(* IEC 61131-3 sources: linesight/plc/src, 5 files *)

(* ---- E_PackML.st ---- *)
// DUT (Enumeration). Numery stanów zgodne z PackML (ISA-TR88.00.02, PackTag Status.StateCurrent).
// Podzbiór: bez stanów przejściowych Holding/Unholding/Suspending/Unsuspending i bez Completing/Complete.
{attribute 'qualified_only'}
TYPE E_PackML :
(
    Clearing  := 1,
    Stopped   := 2,
    Starting  := 3,
    Idle      := 4,
    Suspended := 5,   // przyczyna zewnętrzna: brak produktu na wejściu
    Execute   := 6,
    Stopping  := 7,
    Aborting  := 8,
    Aborted   := 9,
    Held      := 11,  // przyczyna wewnętrzna: zator w maszynie
    Resetting := 15
) INT;
END_TYPE

(* ---- GVL_Line.st ---- *)
// GVL: interfejs linii – wszystko, co wystawiamy przez OPC UA (E3-04).
{attribute 'qualified_only'}
VAR_GLOBAL
    // --- Komendy operatora (zbocze narastające; odpowiednik PackTag Command.CntrlCmd) ---
    xCmdReset     : BOOL;   // Stopped -> Resetting -> Idle
    xCmdStart     : BOOL;   // Idle -> Starting -> Execute
    xCmdStop      : BOOL;   // Idle/Execute/Held/Suspended -> Stopping -> Stopped
    xCmdAbort     : BOOL;   // dowolny stan -> Aborting -> Aborted (wyłącznik awaryjny)
    xCmdClear     : BOOL;   // Aborted -> Clearing -> Stopped

    // --- Wstrzykiwanie awarii (poziom: TRUE = usterka trwa) ---
    xInjJam       : BOOL;   // zator                 -> Held,      iStopReason 101
    xInjNoProduct : BOOL;   // brak produktu         -> Suspended, iStopReason 201
    xInjFault     : BOOL;   // awaria (np. napęd)    -> Aborted,   iStopReason 301
    xInjSlow      : BOOL;   // degradacja: czas cyklu +40 % (dane do wykrywania anomalii, etap 4)
    xInjWear      : BOOL;   // E4-06: zużycie napędu (łożysko) narasta przez tWearRamp; FALSE = naprawa

    // --- Nastawy ---
    tCycleNominal : TIME := T#1500MS;   // nominalny czas cyklu (1 sztuka)
    tWearRamp     : TIME := T#20M;      // E4-06: czas narastania zużycia napędu do 100 %

    // --- Status (tylko do odczytu dla świata) ---
    iStateCurrent    : INT;     // Status.StateCurrent (numer stanu PackML)
    iStopReason      : INT;     // Admin.StopReason.ID: 0 brak, 1 stop operatora, 101 zator,
                                // 201 brak produktu, 301 awaria, 302 abort operatora
    udiProdProcessed : UDINT;   // Admin.ProdProcessedCount (licznik narastający, nie kasujemy)
    udiCycleTime_ms  : UDINT;   // czas ostatniego cyklu [ms] (symulowany)
    rMachSpeed       : REAL;    // Status.CurMachSpeed [szt./min], 0 poza Execute

    // --- E4-06: napęd taśmy (FB_DriveSim), wartości na sztukę ---
    rTorqueMean_Nm   : REAL;    // średni moment w cyklu
    rTorquePeak_Nm   : REAL;    // szczytowy moment w cyklu
    rCurrent_A       : REAL;    // prąd silnika
    rMotorTemp_C     : REAL;    // temperatura silnika (0,1 °C)
    rSimWear         : REAL;    // zużycie 0..1 – prawda symulacji, tylko do oceny modelu (zaokr. 0,01)
END_VAR

(* ---- F_Gauss.st ---- *)
// FUNCTION F_Gauss – szum o rozkładzie zbliżonym do normalnego (średnia 0, odchylenie 1).
// Suma 4 liczb równomiernych z LCG (centralne twierdzenie graniczne); wystarcza do symulacji pomiaru.
// Ziarno przekazywane przez VAR_IN_OUT – stan generatora trzyma wywołujący blok.
// --- część deklaracji ---
FUNCTION F_Gauss : REAL
VAR_IN_OUT
    udiSeed : UDINT;
END_VAR
VAR
    i : INT;
    rSum : REAL;                     // zmienne funkcji startują od 0 przy każdym wywołaniu; nie „s”: S i R to słowa kluczowe IEC (Set/Reset)
END_VAR

// --- część implementacji ---
FOR i := 1 TO 4 DO
    udiSeed := udiSeed * 1103515245 + 12345;
    rSum := rSum + UDINT_TO_REAL((udiSeed / 65536) MOD 32768) / 32768.0;
END_FOR
F_Gauss := (rSum - 2.0) * 1.7320508;    // suma 4 x U(0,1): średnia 2, wariancja 4/12 -> skalowanie do odchylenia 1

(* ---- FB_DriveSim.st ---- *)
// FUNCTION_BLOCK FB_DriveSim – symulacja napędu taśmy (E4-06): moment, prąd, temperatura, zużycie.
// Wartości na sztukę (jak napęd raportujący parametry cyklu), temperatura liczona ciągle.
//   Moment średni   Tm = 2,0 Nm x (1 + 0,15 x zużycie + zimno) + szum 0,06 Nm x (1 + 1,5 x zużycie)
//                   zimno = 0,12 x (40 °C - T) / 18 °C, w zakresie 0..0,12: zimny smar = większe tarcie,
//                   po każdym dłuższym postoju moment jest wyższy o do 12 % i spada, gdy silnik się nagrzeje
//   Moment szczyt.  Tp = Tm x (1,6 + 0,25 x zużycie)     + szum 0,08 Nm x (1 + 2,0 x zużycie)
//   Prąd            I  = 0,8 A + 1,2 A/Nm x Tm            + szum 0,02 A
//   Temperatura     dT/dt = (22 °C + 2,25 x I^2 - T) / 600 s   (inercja 1. rzędu; I = 0 poza Execute)
// Zużycie (np. łożysko): przy xWear rośnie liniowo 0 -> 1 w czasie tWearRamp, bez xWear = 0 (po naprawie).
// Wczesne zużycie ginie w szumie pojedynczej sztuki, a próg na samym momencie myli zużycie z zimnym startem –
// model, który zna temperaturę i kształt cyklu (szczyt/średnia, rozrzut), ma je odróżnić.
// --- część deklaracji ---
FUNCTION_BLOCK FB_DriveSim
VAR_INPUT
    xRun       : BOOL;                 // linia w Execute (napęd pracuje)
    xCycleDone : BOOL;                 // impuls: koniec sztuki – nowe wartości momentu i prądu
    xWear      : BOOL;                 // wstrzyknięte zużycie
    tWearRamp  : TIME := T#20M;        // czas narastania zużycia do 100 %
END_VAR
VAR_OUTPUT
    rTorqueMean : REAL;                // [Nm]
    rTorquePeak : REAL;                // [Nm]
    rCurrent    : REAL;                // [A]
    rTemp       : REAL := 22.0;        // [°C], zaokrąglone do 0,1 (mniej wiadomości przez OPC UA)
    rWear       : REAL;                // 0..1, prawda symulacji – tylko do oceny modelu
END_VAR
VAR
    udiSeed : UDINT := 987654321;
    tLast   : TIME;
    xInit   : BOOL;
    rDt     : REAL;                    // [s] od poprzedniego wywołania
    rT      : REAL := 22.0;            // temperatura bez zaokrąglenia
    rI      : REAL;
    rTm     : REAL;
    rCold   : REAL;                    // dodatkowe tarcie zimnego napędu, 0..0,12
END_VAR
VAR CONSTANT
    T0     : REAL := 2.0;
    TAMB   : REAL := 22.0;
    K_HEAT : REAL := 2.25;
    TAU_S  : REAL := 600.0;
END_VAR

// --- część implementacji ---
IF NOT xInit THEN
    tLast := TIME();
    xInit := TRUE;
END_IF
rDt := TIME_TO_REAL(TIME() - tLast) / 1000.0;
tLast := TIME();

// zużycie
IF xWear AND tWearRamp > T#0S THEN
    rWear := MIN(1.0, rWear + rDt / (TIME_TO_REAL(tWearRamp) / 1000.0));
ELSE
    rWear := 0.0;
END_IF

// temperatura: inercja pierwszego rzędu (metoda Eulera), grzanie proporcjonalne do I^2
IF xRun THEN rI := rCurrent; ELSE rI := 0.0; END_IF
rT := rT + rDt / TAU_S * (TAMB + K_HEAT * rI * rI - rT);
rTemp := DINT_TO_REAL(TRUNC(rT * 10.0)) / 10.0;

// parametry sztuki
IF xCycleDone THEN
    rCold := LIMIT(0.0, 0.12 * (40.0 - rT) / 18.0, 0.12);
    rTm := T0 * (1.0 + 0.15 * rWear + rCold) + 0.06 * (1.0 + 1.5 * rWear) * F_Gauss(udiSeed);
    rTorqueMean := DINT_TO_REAL(TRUNC(rTm * 1000.0)) / 1000.0;
    rTorquePeak := DINT_TO_REAL(TRUNC((rTm * (1.6 + 0.25 * rWear)
                   + 0.08 * (1.0 + 2.0 * rWear) * F_Gauss(udiSeed)) * 1000.0)) / 1000.0;
    rCurrent := DINT_TO_REAL(TRUNC((0.8 + 1.2 * rTm + 0.02 * F_Gauss(udiSeed)) * 1000.0)) / 1000.0;
END_IF

(* ---- PLC_PRG.st ---- *)
// PROGRAM PLC_PRG – maszyna stanów PackML (podzbiór) + symulacja produkcji.
// --- część deklaracji ---
PROGRAM PLC_PRG
VAR
    eState    : E_PackML := E_PackML.Stopped;
    ePrev     : E_PackML := E_PackML.Stopped;
    xNewState : BOOL;
    tonAct    : TON;                 // czas trwania stanów przejściowych (Starting, Stopping, ...)
    tonCycle  : TON;                 // czas cyklu jednej sztuki
    rtReset, rtStart, rtStop, rtAbort, rtClear : R_TRIG;
    tCycle    : TIME := T#1500MS;    // czas bieżącego cyklu (nominalny ± rozrzut)
    udiBase   : UDINT;
    udiSeed   : UDINT := 12345;      // generator pseudolosowy (LCG) do rozrzutu czasu cyklu
    xRun, xRunPrev : BOOL;
    tStart, tNow   : TIME;           // TIME() = czas od startu sterownika; z niego mierzymy rzeczywisty cykl
    xPiece    : BOOL;                // E4-06: impuls – w tym cyklu zadania skończyła się sztuka
    fbDrive   : FB_DriveSim;         // E4-06: symulacja napędu taśmy
END_VAR
VAR CONSTANT
    T_ACT : TIME := T#1S;            // ile trwa każdy stan przejściowy
END_VAR

// --- część implementacji ---
rtReset(CLK := GVL_Line.xCmdReset);
rtStart(CLK := GVL_Line.xCmdStart);
rtStop(CLK := GVL_Line.xCmdStop);
rtAbort(CLK := GVL_Line.xCmdAbort);
rtClear(CLK := GVL_Line.xCmdClear);

// Zegar stanu przejściowego: zeruje się w cyklu, w którym stan się zmienił
xNewState := eState <> ePrev;
ePrev := eState;
tonAct(IN := NOT xNewState, PT := T_ACT);

// Abort ma pierwszeństwo przed wszystkim (jak w PackML: z każdego stanu)
IF (rtAbort.Q OR GVL_Line.xInjFault)
   AND eState <> E_PackML.Aborting AND eState <> E_PackML.Aborted AND eState <> E_PackML.Clearing THEN
    IF GVL_Line.xInjFault THEN
        GVL_Line.iStopReason := 301;
    ELSE
        GVL_Line.iStopReason := 302;
    END_IF
    eState := E_PackML.Aborting;
// Stop operatora z każdego stanu „roboczego”
ELSIF rtStop.Q AND (eState = E_PackML.Idle OR eState = E_PackML.Execute
                    OR eState = E_PackML.Held OR eState = E_PackML.Suspended) THEN
    GVL_Line.iStopReason := 1;
    eState := E_PackML.Stopping;
ELSE
    CASE eState OF
        E_PackML.Stopped:
            IF rtReset.Q THEN eState := E_PackML.Resetting; END_IF

        E_PackML.Resetting:
            GVL_Line.iStopReason := 0;
            IF tonAct.Q THEN eState := E_PackML.Idle; END_IF

        E_PackML.Idle:
            IF rtStart.Q THEN eState := E_PackML.Starting; END_IF

        E_PackML.Starting:
            IF tonAct.Q THEN eState := E_PackML.Execute; END_IF

        E_PackML.Execute:
            IF GVL_Line.xInjJam THEN
                GVL_Line.iStopReason := 101;
                eState := E_PackML.Held;
            ELSIF GVL_Line.xInjNoProduct THEN
                GVL_Line.iStopReason := 201;
                eState := E_PackML.Suspended;
            END_IF

        E_PackML.Held:        // zator usunięty -> wracamy do pracy
            IF NOT GVL_Line.xInjJam THEN
                GVL_Line.iStopReason := 0;
                eState := E_PackML.Execute;
            END_IF

        E_PackML.Suspended:   // produkt wrócił -> wracamy do pracy
            IF NOT GVL_Line.xInjNoProduct THEN
                GVL_Line.iStopReason := 0;
                eState := E_PackML.Execute;
            END_IF

        E_PackML.Stopping:
            IF tonAct.Q THEN eState := E_PackML.Stopped; END_IF

        E_PackML.Aborting:
            IF tonAct.Q THEN eState := E_PackML.Aborted; END_IF

        E_PackML.Aborted:     // kasowanie możliwe dopiero po usunięciu awarii
            IF rtClear.Q AND NOT GVL_Line.xInjFault THEN eState := E_PackML.Clearing; END_IF

        E_PackML.Clearing:
            IF tonAct.Q THEN
                GVL_Line.iStopReason := 0;
                eState := E_PackML.Stopped;
            END_IF
    END_CASE
END_IF

// --- Symulacja produkcji: w Execute jedna sztuka co tCycle ---
// udiCycleTime_ms to ZMIERZONY czas od poprzedniej sztuki (TIME()), a nie zadany tCycle:
// timer widzi czas tylko co cykl zadania, więc rzeczywisty cykl jest dłuższy od zadanego.
xRun := eState = E_PackML.Execute;
IF xRun AND NOT xRunPrev THEN
    tStart := TIME();                // wejście w Execute: liczymy od nowa (postój nie wlicza się do cyklu)
END_IF
xRunPrev := xRun;
tonCycle(IN := xRun, PT := tCycle);
xPiece := tonCycle.Q;
IF tonCycle.Q THEN
    tNow := TIME();
    GVL_Line.udiProdProcessed := GVL_Line.udiProdProcessed + 1;
    GVL_Line.udiCycleTime_ms := TIME_TO_UDINT(tNow - tStart);
    tStart := tNow;
    tonCycle(IN := FALSE);           // kasowanie timera; nowy cykl rusza w następnym cyklu zadania

    // czas następnego cyklu: nominalny (x1,4 przy degradacji) z rozrzutem ±100 ms
    udiBase := TIME_TO_UDINT(GVL_Line.tCycleNominal);
    IF GVL_Line.xInjSlow THEN udiBase := udiBase * 14 / 10; END_IF
    IF udiBase < 300 THEN udiBase := 300; END_IF
    udiSeed := udiSeed * 1103515245 + 12345;
    tCycle := UDINT_TO_TIME(udiBase + (udiSeed / 65536) MOD 201 - 100);
END_IF

// --- E4-06: napęd taśmy ---
fbDrive(xRun := xRun, xCycleDone := xPiece, xWear := GVL_Line.xInjWear, tWearRamp := GVL_Line.tWearRamp);
GVL_Line.rTorqueMean_Nm := fbDrive.rTorqueMean;
GVL_Line.rTorquePeak_Nm := fbDrive.rTorquePeak;
GVL_Line.rCurrent_A     := fbDrive.rCurrent;
GVL_Line.rMotorTemp_C   := fbDrive.rTemp;
GVL_Line.rSimWear       := DINT_TO_REAL(TRUNC(fbDrive.rWear * 100.0)) / 100.0;

// --- Status na zewnątrz ---
GVL_Line.iStateCurrent := eState;
IF eState = E_PackML.Execute AND GVL_Line.udiCycleTime_ms > 0 THEN
    GVL_Line.rMachSpeed := 60000.0 / UDINT_TO_REAL(GVL_Line.udiCycleTime_ms);
ELSE
    GVL_Line.rMachSpeed := 0.0;
END_IF
